FUNCTION_BLOCK fbLightCmdSourceSwitch IMPLEMENTS iLightCmdSource
VAR_INPUT
    LightSwitchState : stSwitchState;
	LightState : stLightState;
END_VAR

{warning 'Add method implementation '}
METHOD Process
VAR_IN_OUT
	CmdEvent	: stLightCmdEvent;
END_VAR

// Exit if switch is idle
IF LightSwitchState.StateType = eSwitchStateType.IDLE THEN
    RETURN;
END_IF

// Short click -> Toggle Light On/Off
IF LightSwitchState.StateType = eSwitchStateType.SHORT_CLICK THEN
	CmdEvent.TargetState.On := NOT LightState.On;
END_IF



CmdEvent.Execute := TRUE;
CmdEvent.Source := eLightCmdSource.SWITCH;
END_METHOD

END_FUNCTION_BLOCK

(* stored: Version 1.1.0.1
   POU fbLightCmdSourceSwitch: Id {bc181d62-640f-4c09-87eb-270fda66e5c5}, SpecialFunc None
   Method Process: Id {761c8d2f-dff1-4a45-bbb9-75d87bb337f7} *)
